(* IEC 61131-3 sources: PLC-Static-Analysis/modules/plc-rules/src/test/resources/PLCA-Q015/custom, 1 file *)

(* ---- c.st ---- *)
FUNCTION_BLOCK FB_Valve
VAR_INPUT
    xOpen : BOOL;
    bClose : BOOL; // PLCA-Q015
END_VAR
END_FUNCTION_BLOCK
